TYPE ST_PatchFeedStatus :
STRUCT
    bPermitted : BOOL;
    bConfigured : BOOL;
    bWasteRollDemand : BOOL;
    bBusy : BOOL;
    bFault : BOOL;
    bResetPending : BOOL;
    udiErrorId : UDINT;
    sDiagnostic : STRING(160);
    bPatchFeedRollDemand : BOOL;
    bDriveBusy : BOOL;
    bDriveRunDemand : BOOL;
END_STRUCT
END_TYPE

(* stored: Version 1.1.0.1, ProductVersion 3.1.4026.18
   DUT ST_PatchFeedStatus: Id {7dc67d44-8589-4f59-acf6-74dda7d36fdc} *)
